// Core S3.12 - the SET target in engineering units, latched at Execute.
TYPE ST_AnalogOutputParCmd :
STRUCT
    Target : LREAL;
END_STRUCT
END_TYPE

(* stored: Version 1.1.0.1, ProductVersion 3.1.4024.12
   DUT ST_AnalogOutputParCmd: Id {161eb2ca-8da9-4da3-bd38-5a121ba0add4} *)
